FUNCTION_BLOCK INT2UINT (* Writing INT from input to UINT output *)
  (* Standard: 61499-1 *)
  (* Version 1.0, 2023-03-07, Bianca Wiesmayr *)
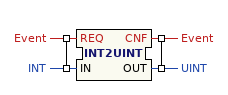
  EVENT_INPUT
    REQ WITH IN; (* Normal Execution Request *)
  END_EVENT
  EVENT_OUTPUT
    CNF WITH OUT; (* Execution Confirmation *)
  END_EVENT
  VAR_INPUT
    IN : INT;
  END_VAR
  VAR_OUTPUT
    OUT : UINT;
  END_VAR
  ALGORITHM REQ IN ST:
	OUT:=INT_TO_UINT(IN);
  END_ALGORITHM
END_FUNCTION_BLOCK
